{attribute 'qualified_only'}
VAR_GLOBAL
	// Komutlar (ADS schreibt, FB_Kessel verarbeitet)
	CmdHeizung : BOOL;
	CmdPumpe : BOOL := TRUE;
	CmdSollwert : LREAL := 60.0;
	CmdNotaus : BOOL;
	CmdNotausReset : BOOL;

	// Zustand (ADS liest, nur PLC schreibt)
	Temperatur : LREAL := 20.0;
	Heizung : BOOL;
	Pumpe : BOOL := TRUE;
	Sollwert : LREAL := 60.0;
	Notaus : BOOL;
	ZielAlarmSekunden : LREAL;
	AutoGestoppt : BOOL;
END_VAR

(* stored: Version 1.1.0.1, ProductVersion 3.1.4024.32
   GVL GVL: Id {5D4EAF60-7182-4D9E-BFA0-2B3C4D5E6F70} *)
